TYPE eShutterCmdSource :
(
    NONE,
    SWITCH,
    HA,
    SCHEDULER,
	ROOM
);
END_TYPE

(* stored: Version 1.1.0.1
   DUT eShutterCmdSource: Id {e1d68600-0f36-4136-8459-342dec891c86} *)
